// TIA Portal V20 export
// export: Created 2026-10-19T18:04:21.7743256Z, ExportSetting WithDefaults, DisplayName Totally Integrated Automation Portal, DisplayVersion V20 Update 6, DisplayName TIA Portal Openness, DisplayVersion V20 Update 6, DisplayName TIA Portal Version Control Interface, DisplayVersion V20 Update 6, DisplayName SINAMICS Startdrive Advanced, DisplayVersion V20 SP1, DisplayName SINAMICS Startdrive G130, G150, S120, S150, SINAMICS MV, G220, S200, S210, DisplayVersion V20 SP1, DisplayName SINAMICS Startdrive G110M, G120, G120C, G120D, G120P, G115D, DisplayVersion V20 SP1, DisplayName STEP 7 Professional, DisplayVersion V20 Update 6, DisplayName STEP 7 Safety, DisplayVersion V20 Update 2, DisplayName WinCC Basic/Comfort/Advanced, DisplayVersion V20 Update 6, DisplayName WinCC Unified, DisplayVersion V20 Update 6
FUNCTION_BLOCK "Safety_Stops_FB"   // FB7, SCL
{ S7_Optimized_Access := 'TRUE' }
VERSION : 0.1
// stored: AutoNumber true, IsIECCheckEnabled false, IsRetainMemResEnabled false, MemoryReserve 100, SetENOAutomatically false, UDAEnableTagReadback false
   VAR_INPUT
      Mode : UInt;
      Timeout : UInt;
      Reset : Bool;
      Up : Bool;
      Down : Bool;
   END_VAR
   VAR_OUTPUT
      Rotate : Bool;
   END_VAR
   VAR_IN_OUT
      Sfts_Control : "Sfts_Control";
   END_VAR
   VAR
      State : UInt;
      LP_Timer { ExternalAccessible := 'False'; ExternalVisible := 'False'; ExternalWritable := 'False'} : TON_TIME;
      IEC_Timer_0_Instance { S7_SetPoint := 'True'} : TOF_TIME;
      Timer_1 : Time;
   END_VAR
BEGIN
   #Sfts_Control.Enabled := #Sfts_Control.Instruction.Enable := #Mode = 2 OR #Mode = 3;

   //MODES
   IF (#Mode = 1 OR #Mode = 5) AND NOT #Sfts_Control.Error THEN
       #State := 500;
   END_IF;

   (*
   TODO
   1. Need to add the mode and running checks for manual mode
   2. Add output for safety stop brake.

   Mode select is done via the HMI. Might add external mode select switches.

           Mode select mask:
           0: Disabled
           1: Manual
           2: Semi-Auto
           3: Auto
           4: Teach - N/A for Cnv
           5: Maintenance

   Device ID Format: XXYYZZ    
   XX = Device type   
       01   VTD
       10  Cnv_Front_of_VTD
       11  Cnv_Rear_of_VTD
       12  Cnv_On_Extractor
       20  Safety_Stop_Front_of_VTD
       21  Safety_Stop_Rear_of_VTD
   YY = Floor   
   ZZ = VTD Connected to 
   *)

   REGION Assign Inputs
       #Sfts_Control.Inputs.LP_Extended := #Up;
       #Sfts_Control.Inputs.LP_Retracted := #Down;
   END_REGION

   REGION Cyclic Checks
       //Update variables
       #Sfts_Control.SM_State := #State;

       #LP_Timer(IN := #Sfts_Control.Running,
                 PT := UINT_TO_TIME(#Timeout));

       //STOPPER STATE
       IF #Sfts_Control.Inputs.LP_Extended AND NOT #Sfts_Control.Inputs.LP_Retracted THEN
           #Sfts_Control.LP_State := 1; // EXTENDED
       ELSIF NOT #Sfts_Control.Inputs.LP_Extended AND #Sfts_Control.Inputs.LP_Retracted THEN
           #Sfts_Control.LP_State := 0; //RETRACTED
       ELSE
           #Sfts_Control.LP_State := 2; //LOST
       END_IF;;
   END_REGION

   REGION Auto Mode

           CASE #State OF
               0: //IDLE MODE
                   IF #Mode = 2 OR #Mode = 3 THEN
                       IF #Sfts_Control.Instruction.Enable AND #Sfts_Control.Error = 0 THEN
                           #Sfts_Control.Enabled := TRUE;
                           #State := 10;
                       END_IF;
                   END_IF;
               10: //Standby
                   IF NOT #Sfts_Control.Running AND #Sfts_Control.Error = 0 AND #Sfts_Control.Instruction.LP_Extend THEN
                       IF #Sfts_Control.Inputs.LP_Extended THEN
                           ; // Complete the task as the LP ar already extended
                       ELSIF #Sfts_Control.Inputs.LP_Retracted THEN
                           #Sfts_Control.Running := True;
                           #State := 20;
                       ELSE
                           #Sfts_Control.Error := 0; //Unknown locking pin state
                           #State := 400;
                       END_IF;
                   ELSIF NOT #Sfts_Control.Running AND #Sfts_Control.Error = 0 AND #Sfts_Control.Instruction.LP_Retract THEN
                       IF #Sfts_Control.Inputs.LP_Retracted THEN
                           ; // Complete the task as the LP ar already extended
                       ELSIF #Sfts_Control.Inputs.LP_Extended THEN
                           #Sfts_Control.Running := True;
                           #State := 40;
                       ELSE
                           #Sfts_Control.Error := 0; //Unknown locking pin state
                           #State := 400;
                       END_IF;
                   END_IF;

               20: //Extend safety locking pins
                   #Sfts_Control.Motor_Extend := TRUE;
                   IF #Sfts_Control.Inputs.LP_Extended THEN
                       #Sfts_Control.Motor_Extend := FALSE;
                       #Sfts_Control.Running := FALSE;
                       #State := 0;
                   END_IF;

               40: //Retract safety locking pins
                   #Sfts_Control.Motor_Retract := TRUE;
                   IF #Sfts_Control.Inputs.LP_Retracted THEN
                       #Sfts_Control.Motor_Retract := FALSE;
                       #Sfts_Control.Running := FALSE;
                       #State := 0;
                   END_IF;

               400: // Error#Sfts_Control
                   #Sfts_Control.Motor_Retract := FALSE;
                   #Sfts_Control.Motor_Extend := FALSE;
                   #Sfts_Control.Running := FALSE;
                   #LP_Timer(IN := FALSE,
                             PT := T#0S);
                   IF #Reset THEN
                       #Sfts_Control.Error := FALSE;
                       #State := 0;
                   END_IF;

               500:
                   IF #Sfts_Control.Instruction.Manual_Extend AND NOT #Sfts_Control.Inputs.LP_Extended THEN
                       #Sfts_Control.Motor_Extend := TRUE;
                       #Sfts_Control.Running := TRUE;
                   ELSIF #Sfts_Control.Instruction.Manual_Retract AND NOT #Sfts_Control.Inputs.LP_Retracted THEN
                       #Sfts_Control.Motor_Retract := TRUE;
                       #Sfts_Control.Running := TRUE;
                   ELSE
                       #Sfts_Control.Motor_Extend := FALSE;
                       #Sfts_Control.Motor_Retract := FALSE;
                       #Sfts_Control.Running := FALSE;
                   END_IF;

                   IF #Mode <> 1 AND #Mode <> 5 THEN
                       #State := 0;
                   END_IF;
           END_CASE;
   END_REGION

   REGION Cyclic Error Checks
       IF #Sfts_Control.Inputs.LP_Extended AND #Sfts_Control.Inputs.LP_Retracted THEN
           #Sfts_Control.Error := TRUE; //Cant have the locking pins extended and retracted at the same time11
       END_IF;

       // Statement section REGION
       IF #LP_Timer.Q THEN
           #Sfts_Control.Error := TRUE;//locking pin timeout
       END_IF;

       IF #Sfts_Control.Error THEN
           #State := 400;
       END_IF;
   END_REGION

   REGION Assign outputs
       #IEC_Timer_0_Instance(IN := #Sfts_Control.Motor_Extend OR #Sfts_Control.Motor_Retract,
                             PT := #Timer_1,
                             Q => #Rotate);
   END_REGION
END_FUNCTION_BLOCK
